(* IEC 61131-3 sources: daoli-st-library/DL_MathData (part 32) *)

(* ---- FC_DL_RangeOverlapCheck.st ---- *)
(*==============================================================================
 * 组件名称 (Component)  : FC_DL_RangeOverlapCheck
 * 所属子库 (Sublibrary) : DL_MathData
 * 当前版本 (Version)    : 1.0.0
 * 分类     (Category)   : 区间关系判定函数（Function · Comparator / Pure function）
 * 兼容性   (Platform)   : CODESYS 3.5 / TwinCAT 3 / 汇川 InoProShop / Machine Expert
 *                         仅依赖 Standard.library（ABS / MIN / MAX），零厂商方言
 * 功能描述 (Function)   : 判定两个实数区间 A、B 的几何关系（相离 / 仅端点相接 /
 *                         部分重叠 / 一方包含另一方 / 完全相等），并输出重叠长度。
 *                         输入是 4 个端点而非 1 个测量值，返回值为关系枚举，全程
 *                         无内部状态，可任意频次调用。用于配方参数域校验、时间窗
 *                         互斥检查、公差带叠加分析、安全包络与工艺窗口对撞检查。
 *
 * 【引脚契约 / Pin contract】
 *   输入 fA1        : REAL — 区间 A 端点 1 [任意工程单位]，无序自动对调；
 *   输入 fA2        : REAL — 区间 A 端点 2，同上；
 *   输入 fB1        : REAL — 区间 B 端点 1，无序自动对调；
 *   输入 fB2        : REAL — 区间 B 端点 2，同上；
 *   输入 bIncA      : BOOL — A 是否闭区间（含端点），默认 TRUE；
 *   输入 bIncB      : BOOL — B 是否闭区间，默认 TRUE；
 *   输出 fOverlapSpan : REAL — 重叠长度 [与输入同单位]，无重叠 = 0.0，恒非负；
 *   输出 bTouching    : BOOL — 仅端点相接（重叠长度 0 但边界重合）；
 *   输出 bValid       : BOOL — 四个输入全部有限（非 NaN、非无穷）= TRUE；
 *   输出 uErrorId     : UDINT — 事件码，0 = 无。本件全部码为信息级。
 *   返回  值          : E_DL_RangeRelation — 区间关系枚举，见下方成员语义表。
 *
 * 【关系枚举语义 / Relation enum semantics（同文件发布）】
 *   eInvalid  = 0  — 输入含非有限值（NaN / 无穷），关系不可判，重叠长度 0.0；
 *   eDisjoint = 10 — 完全相离（两区间之间有正间隙）；
 *   eTouching = 20 — 仅端点相接，重叠长度 0.0，bTouching 置位；
 *   ePartial  = 30 — 部分重叠（互相不包含，重叠长度大于 0）；
 *   eContains = 40 — 一方包含另一方（含端点恰好重合的包含）；
 *   eEqual    = 50 — 两端点均在容差内相等，重叠长度 = 区间长度。
 *
 * 【判定次序 / Decision order（写死，避免多解）】
 *   ① 有限性闸门 → 全部有限才继续，否则返回 eInvalid 并置 0121；
 *   ② 端点归一 → 每个区间内部排序，保证「下限 <= 上限」；
 *   ③ 相等判定 → 两端点同时落在容差内即 eEqual（先判，避免被包含分支吞掉）；
 *   ④ 相离判定 → 任一侧上限严格小于对侧下限减去容差，即 eDisjoint；
 *   ⑤ 相接判定 → 任一侧上限与对侧下限重合（容差内），即 eTouching；
 *   ⑥ 包含判定 → 一侧下限不大于对侧下限且上限不小于对侧上限，即 eContains；
 *   ⑦ 其余 → ePartial（此时重叠长度必然大于 0，无需再判）。
 *   次序不可调换：相等必须先于包含，相离必须先于相接，相接必须先于部分重叠。
 *
 * 【开闭区间口径 / Open and closed intervals（防误解声明）】
 *   ① 几何关系与开闭无关：「相接」只描述两组端点几何重合，开区间同样判相接；
 *   ② 开闭只影响「相接处那一个点是否属于公共交集」，其判据为
 *      bTouching AND bIncA AND bIncB —— 调用方按此合成，本件不额外输出第三态；
 *   ③ 部分重叠与包含的重叠长度按端点差值计算，不做「开区间减去两个端点」的
 *      离散化折算：连续量工程口径下端点测度为零，减去端点会引入 1 个单位误差；
 *   ④ 相等判定用容差而非判等（浮点判等红线）：两端点差值绝对值均小于容差即认为
 *      相等，容差取 1.0E-6，对应工程上「不可分辨」的量级。
 *
 * 【数值安全 / Numeric safety】
 *   N1 非有限值用「区间比较取反」识别：NaN 参与任何有序比较均为假，
 *      故 NOT(下限比较 AND 上限比较) 同时覆盖 NaN 与正负无穷，无需判等；
 *   N2 重叠长度在返回前置零下限保护：极少数退化输入可能算出负零附近的微小负值，
 *      一律钳到 0.0，保证输出恒非负（下游可直接做累加不打补丁）；
 *   N3 全件无除法、无开方、无累加迭代，不存在除零与溢出风险；
 *   N4 全件无循环、无数组访问，不存在越界风险。
 *
 * 【边界防错清单 / Boundary guard list】
 *   B1 输入非有限 → bValid FALSE、返回 eInvalid、重叠长度 0.0、置 0121（信息级）；
 *   B2 端点无序（如 A = [10, 0]）→ 自动对调后按归一区间判定，不置任何码；
 *   B3 零长度区间（两端点相等）→ 合法输入，参与全部关系判定，不特殊对待；
 *   B4 相接与部分重叠的边界由容差分割：端点差值绝对值小于容差判相接，
 *      否则按下限比较判重叠，容差量级远小于工程分辨率，不会误判真实重叠；
 *   B5 包含判定允许端点恰好重合（A 包含 B 且共端点），此时关系为 eContains
 *      而非 eEqual（eEqual 要求两端点都相等，先判，语义不重叠）。
 *
 * 【与既有件的职责边界 / Family separation（本族唯一二元件）】
 *   FC_DL_LimitClassify    = 判单个测量值落在哪一档（单点 → 档位）；
 *   FC_DL_Hysteresis       = 判单个测量值的迟滞切换（单点 + 历史 → 开关）；
 *   FB_DL_ToleranceWindow  = 判单个测量值是否落在公差带（单点 → 布尔）；
 *   本件                   = 判两个区间之间的关系（四点 → 关系枚举），
 *   输入元数不同、返回类型不同，四者不可互相替代。
 *
 * 【调用示例 / Call example（仅行注释，不嵌套块注释）】
 *   // 配方切换前校验：新工艺窗口与安全包络是否相撞
 *   // eRel := FC_DL_RangeOverlapCheck(fA1 := fSafeLo, fA2 := fSafeHi,
 *   //        fB1 := fNewLo, fB2 := fNewHi, bIncA := TRUE, bIncB := TRUE,
 *   //        fOverlapSpan => fOverlap, bTouching => bTouch,
 *   //        bValid => bCfgValid, uErrorId => uRelErr);
 *   // IF eRel = E_DL_RangeRelation.ePartial OR eRel = E_DL_RangeRelation.eContains THEN
 *   //     bRejectRecipe := TRUE;
 *   // END_IF
 *
 * 【平台移植注意 / Porting notes】
 *   仅用 ABS / MIN / MAX 三个标准函数与有序比较，无舍入模式依赖；
 *   容差与有限性阈值全部来自 VAR CONSTANT，换平台无需改逻辑；
 *   返回枚举类型随本文件发布，导入顺序上本文件不依赖任何其他 DL_ 组件。
 *
 * 【工程背景与应用场景 / Background and use cases】
 *   ① 配方参数域校验：新配方允许的温度带与设备安全包络相撞时拒绝下发；
 *   ② 时间窗互斥检查：两班次的作业窗若部分重叠，提示排程冲突；
 *   ③ 公差带叠加：来料公差带与装配公差带仅端点相接时，判定为「临界合格」；
 *   ④ 安全包络对撞：机器人可达包络与围栏安全距离带的重叠长度用于风险评估。
 *
 * 【验收向量 / Acceptance vectors】
 *   V1 部分重叠：A = [0, 10]、B = [5, 15] → ePartial、重叠长度 5.0；
 *   V2 端点相接：A = [0, 10]、B = [10, 20] → eTouching、重叠长度 0.0、bTouching；
 *   V3 包含：A = [0, 10]、B = [2, 8] → eContains、重叠长度 6.0；
 *   V4 相离：A = [0, 10]、B = [20, 30] → eDisjoint、重叠长度 0.0；
 *   V5 相等：A = [0, 10]、B = [0, 10] → eEqual、重叠长度 10.0；
 *   V6 无序端点：A = [10, 0]、B = [5, 15] → 归一后同 V1，ePartial、5.0；
 *   V7 非有限：fA1 为 NaN → eInvalid、bValid FALSE、uErrorId 0121。
 *
 * 【事件码表 / Event code table（全部信息级，不置报警位）】
 *   16#0001_0121  输入含非有限值，关系不可判，返回 eInvalid 与重叠长度 0.0。
 *
 * 修订历史 (Revision)   :
 *   2026-11-15  v1.0.0  首版落盘（Round 11 · 泳道 A · LGF Comparator 组）
 *
 * 同文件发布类型 (Co-published type) : E_DL_RangeRelation（本函数返回枚举，
 *   按库内惯例随宿主 POU 同文件发布，禁止在其他文件重复声明同名枚举）。
 *============================================================================*)
TYPE E_DL_RangeRelation :
(
    eInvalid  := 0,    // 输入非有限值，关系不可判 / Inputs not finite, relation undecidable
    eDisjoint := 10,   // 完全相离，存在正间隙 / Fully disjoint with a positive gap
    eTouching := 20,   // 仅端点相接，重叠长度为零 / Endpoint touch only, zero overlap
    ePartial  := 30,   // 部分重叠，互不包含 / Partial overlap, neither contains the other
    eContains := 40,   // 一方包含另一方 / One range contains the other
    eEqual    := 50    // 两端点均在容差内相等 / Both endpoints equal within tolerance
);
END_TYPE

FUNCTION FC_DL_RangeOverlapCheck : E_DL_RangeRelation
VAR_INPUT
    fA1     : REAL;                        // 区间 A 端点 1 [工程单位]，无序自动对调 / Range A endpoint 1 [EU], auto-swapped
    fA2     : REAL;                        // 区间 A 端点 2 [工程单位] / Range A endpoint 2 [EU]
    fB1     : REAL;                        // 区间 B 端点 1 [工程单位]，无序自动对调 / Range B endpoint 1 [EU], auto-swapped
    fB2     : REAL;                        // 区间 B 端点 2 [工程单位] / Range B endpoint 2 [EU]
    bIncA   : BOOL := TRUE;                // A 是否闭区间，含端点 / A closed interval flag, endpoints included
    bIncB   : BOOL := TRUE;                // B 是否闭区间，含端点 / B closed interval flag, endpoints included
END_VAR
VAR_OUTPUT
    fOverlapSpan : REAL;                   // 重叠长度 [工程单位]，无重叠 0.0，恒非负 / Overlap length [EU], zero when none, never negative
    bTouching    : BOOL;                   // 仅端点相接（几何重合，与开闭无关）/ Endpoint touch only, independent of openness
    bValid       : BOOL;                   // 四个输入全为有限值 / All four inputs are finite
    uErrorId     : UDINT;                  // 事件码，0 = 无 / Event code, 0 = none
END_VAR
VAR
    _fLoA   : REAL;                        // 区间 A 归一下限 [工程单位] / Normalised lower bound of range A [EU]
    _fHiA   : REAL;                        // 区间 A 归一上限 [工程单位] / Normalised upper bound of range A [EU]
    _fLoB   : REAL;                        // 区间 B 归一下限 [工程单位] / Normalised lower bound of range B [EU]
    _fHiB   : REAL;                        // 区间 B 归一上限 [工程单位] / Normalised upper bound of range B [EU]
    _fTmp   : REAL;                        // 对调临时量 [工程单位] / Swap temporary [EU]
    _fLo    : REAL;                        // 重叠区间下限 = 两个下限的较大者 [工程单位] / Overlap lower bound, the larger of both [EU]
    _fHi    : REAL;                        // 重叠区间上限 = 两个上限的较小者 [工程单位] / Overlap upper bound, the smaller of both [EU]
    _bFinite : BOOL;                       // 有限性闸门标志 / Finiteness gate flag
END_VAR
VAR CONSTANT
    DL_FLOAT_EPS  : REAL  := 1.0E-6;       // 端点比较容差 [工程单位] / Endpoint comparison epsilon [EU]
    DL_INF_LIM    : REAL  := 1.0E37;       // 非有限值判据阈值，超此视为无穷 / Non-finite threshold, beyond is infinity
    DL_SPAN_ZERO  : REAL  := 0.0;          // 重叠长度下界，恒非负 / Overlap length lower bound, never negative
    DL_ERR_NONFIN : UDINT := 16#0001_0121; // 输入非有限值的信息级码 / Info code for non-finite inputs
END_VAR

(*------------------------------------------------------------------------------
 * 段 1｜返回值与输出预置（函数必须先给出安全返回值）
 *      Preset the return value and the outputs
 *   默认返回 eInvalid：任何早退路径都天然带着「不可判」语义，不会误报相离。
 *-----------------------------------------------------------------------------*)
FC_DL_RangeOverlapCheck := E_DL_RangeRelation.eInvalid;   // 返回值预置不可判（Return preset to undecidable）
fOverlapSpan := DL_SPAN_ZERO;              // 重叠长度预置 0（Overlap span preset to zero）
bTouching    := FALSE;                     // 相接标志预置（Touch flag preset）
bValid       := TRUE;                      // 有效性预置通过（Validity preset to pass）
uErrorId     := 16#0000_0000;              // 事件码预清零（Event code preset to zero）
_bFinite     := TRUE;                      // 有限性闸门预置通过（Finiteness gate preset to pass）

(*------------------------------------------------------------------------------
 * 段 2｜有限性闸门（边界 B1 / 数值安全 N1）
 *      Finiteness gate
 *   NaN 与任何有序比较的结果均为假，故「比较区间取反」同时覆盖 NaN 与无穷，
 *   不必使用浮点判等，也不依赖任何厂商的非有限值判定函数。
 *-----------------------------------------------------------------------------*)
IF NOT ((fA1 <= DL_INF_LIM) AND (fA1 >= -DL_INF_LIM)) THEN   // 端点 A1 非有限（A1 not finite）
    _bFinite := FALSE;                     // 闸门关闭（Close the gate）
END_IF
IF NOT ((fA2 <= DL_INF_LIM) AND (fA2 >= -DL_INF_LIM)) THEN   // 端点 A2 非有限（A2 not finite）
    _bFinite := FALSE;                     // 闸门关闭（Close the gate）
END_IF
IF NOT ((fB1 <= DL_INF_LIM) AND (fB1 >= -DL_INF_LIM)) THEN   // 端点 B1 非有限（B1 not finite）
    _bFinite := FALSE;                     // 闸门关闭（Close the gate）
END_IF
IF NOT ((fB2 <= DL_INF_LIM) AND (fB2 >= -DL_INF_LIM)) THEN   // 端点 B2 非有限（B2 not finite）
    _bFinite := FALSE;                     // 闸门关闭（Close the gate）
END_IF

IF NOT _bFinite THEN                       // 任一输入不可判（Any input undecidable）
    bValid   := FALSE;                     // 有效性置假（Validity cleared）
    uErrorId := DL_ERR_NONFIN;             // 置非有限值信息码（Raise the non-finite info code）
    RETURN;                                // 早退，返回值保持 eInvalid（Early exit, return stays eInvalid）
END_IF

(*------------------------------------------------------------------------------
 * 段 3｜端点归一（边界 B2：无序端点自动对调）
 *      Endpoint normalisation, unordered endpoints are swapped
 *   归一后不可能出现「下限大于上限」，后续全部比较都是同向比较。
 *-----------------------------------------------------------------------------*)
_fLoA := fA1;                              // A 下限暂存端点 1（A lower bound takes endpoint 1）
_fHiA := fA2;                              // A 上限暂存端点 2（A upper bound takes endpoint 2）
IF _fLoA > _fHiA THEN                      // 端点逆序（Endpoints in reverse order）
    _fTmp := _fLoA;                        // 暂存下限（Save the lower bound）
    _fLoA := _fHiA;                        // 下限取原上限（Lower takes the former upper）
    _fHiA := _fTmp;                        // 上限取原下限（Upper takes the former lower）
END_IF

_fLoB := fB1;                              // B 下限暂存端点 1（B lower bound takes endpoint 1）
_fHiB := fB2;                              // B 上限暂存端点 2（B upper bound takes endpoint 2）
IF _fLoB > _fHiB THEN                      // 端点逆序（Endpoints in reverse order）
    _fTmp := _fLoB;                        // 暂存下限（Save the lower bound）
    _fLoB := _fHiB;                        // 下限取原上限（Lower takes the former upper）
    _fHiB := _fTmp;                        // 上限取原下限（Upper takes the former lower）
END_IF

_fLo := MAX(_fLoA, _fLoB);                 // 重叠下限 = 两个下限的较大者（Overlap lower bound）
_fHi := MIN(_fHiA, _fHiB);                 // 重叠上限 = 两个上限的较小者（Overlap upper bound）

(*------------------------------------------------------------------------------
 * 段 4｜关系判定（判定次序写死：相等 → 相离 → 相接 → 包含 → 部分）
 *      Relation decision in the frozen order
 *   次序不可调换，理由见头注释「判定次序」段；每支都显式给出重叠长度。
 *-----------------------------------------------------------------------------*)
IF (ABS(_fHiA - _fHiB) < DL_FLOAT_EPS) AND (ABS(_fLoA - _fLoB) < DL_FLOAT_EPS) THEN
    FC_DL_RangeOverlapCheck := E_DL_RangeRelation.eEqual;   // 相等：两端点均在容差内（Both endpoints equal within epsilon）
    fOverlapSpan := _fHiA - _fLoA;         // 重叠长度 = 区间长度（Overlap equals the range length）
ELSIF (_fHiA < _fLoB - DL_FLOAT_EPS) OR (_fHiB < _fLoA - DL_FLOAT_EPS) THEN
    FC_DL_RangeOverlapCheck := E_DL_RangeRelation.eDisjoint; // 相离：存在正间隙（A positive gap exists）
    fOverlapSpan := DL_SPAN_ZERO;          // 相离无重叠（No overlap when disjoint）
ELSIF (ABS(_fHiA - _fLoB) < DL_FLOAT_EPS) OR (ABS(_fHiB - _fLoA) < DL_FLOAT_EPS) THEN
    FC_DL_RangeOverlapCheck := E_DL_RangeRelation.eTouching; // 相接：端点几何重合（Endpoints coincide geometrically）
    fOverlapSpan := DL_SPAN_ZERO;          // 相接重叠长度为零（Zero overlap on a touch）
    bTouching    := TRUE;                  // 置相接标志（Raise the touch flag）
ELSIF ((_fLoA <= _fLoB + DL_FLOAT_EPS) AND (_fHiA >= _fHiB - DL_FLOAT_EPS)) OR
      ((_fLoB <= _fLoA + DL_FLOAT_EPS) AND (_fHiB >= _fHiA - DL_FLOAT_EPS)) THEN
    FC_DL_RangeOverlapCheck := E_DL_RangeRelation.eContains; // 包含：一方完全覆盖另一方（One range covers the other）
    fOverlapSpan := _fHi - _fLo;           // 重叠长度 = 被包含区间的长度（Overlap equals the inner range length）
ELSE
    FC_DL_RangeOverlapCheck := E_DL_RangeRelation.ePartial; // 部分重叠：互不包含（Partial overlap, neither contains）
    fOverlapSpan := _fHi - _fLo;           // 重叠长度 = 交集长度（Overlap equals the intersection length）
END_IF

(*------------------------------------------------------------------------------
 * 段 5｜重叠长度非负保护（数值安全 N2）
 *      Non-negative guard of the overlap span
 *   浮点舍入可能让理论为零的交集算出极小的负值，一律钳到 0，
 *   保证下游可直接累加与比较，不必各自打补丁。
 *-----------------------------------------------------------------------------*)
IF fOverlapSpan < DL_SPAN_ZERO THEN        // 重叠长度出现负值（A negative span appeared）
    fOverlapSpan := DL_SPAN_ZERO;          // 钳到 0，维持非负承诺（Clamp to zero, keep the promise）
END_IF
END_FUNCTION

(* ---- FC_DL_StringFixedField.st ---- *)
(*==============================================================================
 * 组件名称 (Component)  : FC_DL_StringFixedField
 * 所属子库 (Sublibrary) : DL_MathData
 * 归属目录 (Directory)  : C:\Library\DL_MathData
 * 当前版本 (Version)    : 1.0.0
 * 分类/来源标签         : 函数（FUNCTION）· 纯函数 · 定宽字段填充与对齐
 *                         lgf-datahandling / fixed-field / r37-reference
 * 兼容性   (Platform)   : CODESYS 3.5 / TwinCAT 3 / 汇川 InoProShop / 施耐德
 *                         Machine Expert；仅用 Standard.library 的 LEN / MID /
 *                         CONCAT / MIN，字符串声明一律显式带长度
 * 功能一句话 (Summary)  : 把任意文本装进定宽字段（左对齐或右对齐、指定填充字符），
 *                         并在发生裁剪时显式置截断标志与事件码。
 *
 * 本件存在的意义 (Why this unit exists)：
 *   本件存在的意义是把 R37 变成可复制的写法。全库所有「往定长缓冲写串」的地方，
 *   都可以照本件的四步顺序抄：先算一次源长度，再与目标宽度比较，比较成立就先置
 *   截断标志与码，最后才写缓冲。顺序一旦颠倒（先 CONCAT 再回夹、或回夹时不置标志），
 *   现场就会出现「字段看着对、内容被砍了一半、日志里一个字都没有」的事故。
 *   本件是全库唯一一处必须在写入前预判长度的地方，因此写成了可当范本读的样子。
 *
 * 功能描述 (Function)   : 先校验宽度契约，再解析填充字符，然后一次取源长度并与宽度
 *                         比较，按允许与否决定「截断写出」或「拒绝构造」，最后用
 *                         CONCAT 把核心段与填充段拼成恰好 nWidth 个字符的字段。
 *                         典型现场用途：定长报文拼装（固定列宽协议）、CSV 列对齐、
 *                         HMI 固定列显示、条形码定长补位、打印模板的等宽排版。
 * 与既有件边界 (Boundary): FC_DL_StringTrim 去首尾空白、FC_DL_StringSplit 拆分、
 *                         FC_DL_StringReplaceAll 替换。三者都改变内容而不改宽度；
 *                         本件只改宽度与对齐，内容字符顺序不动（除裁剪尾部）。
 *                         宽度是契约参数，本件不猜、不钳、不补零。
 * 设计要点 (Key notes)  : ① 源长度只取一次（R38），其后所有比较与循环上界都用该副本；
 *                         ② 裁剪判定先于任何写入（R37），标志置位先于结果构造；
 *                         ③ 拼装只用 CONCAT 与单字符填充，绝不用取子串的函数去「凑宽度」，
 *                           也不做「先拼后夹」的回夹写法；
 *                         ④ 出口长度天然等于宽度（核心段加填充段恰好补齐），总长不超过
 *                           声明上限，故不存在赋值时的静默截断；
 *                         ⑤ 每次进入先把结果清空，杜绝上一次调用的残留字符。
 *                         ⑥ 纯函数：无内部状态、无跨周期残留，同入参同结果。
 *
 * 【R37 四步顺序（本件样板，调用方照抄即可）】
 *   第 1 步  nSrcLen := LEN(sValue)                         只取一次，锁存
 *   第 2 步  IF nSrcLen > MIN(nWidth, DL_SFF_MAXLEN) THEN  与目标宽度比较（宽度与上限取小）
 *   第 3 步      bTruncated := TRUE                          先置标志，先于任何写入
 *   第 4 步      按 bAllowTrunc 决定截断写出还是拒绝构造     最后才写缓冲
 *
 * 【验收向量 / Acceptance vectors】
 *   V1  源「ABC」、宽度 6、左对齐 → 字段「ABC 加三个空格」、写出 6、不截断
 *   V2  源「ABC」、宽度 6、右对齐 → 字段「三个空格加 ABC」、写出 6
 *   V3  V-B 主向量（R37 核心）：源「ABCDEFGHIJ」、宽度 5、允许截断
 *       → 字段「ABCDE」、截断标志为真、码 0147；裁剪发生必须有人报警
 *   V4  V-B 拒绝路：同源同宽、不允许截断 → 返回假、字段空串、写出 0、码 0148、
 *       截断标志仍为真（事实发生了，只是没写出去）
 *   V5  V-A 域外：宽度 0 或宽度 300 → 返回假、码 0224；宽度不钳位，
 *       因为宽度是契约，猜不得
 *   V6  残留专测：连续两次调用，第二次源为空串 → 字段必须是纯填充，不残留上次内容
 *   V7  V-D 填充字符纠正：填充串为空 → 退回空格并置 0149，字段仍按宽度构造
 *
 * 开源溯源 (Origin)     : 来源标签 lgf-datahandling。LGF（Libre Graphical Framework）
 *                         为免费闭源发布的公开函数库手册，本件仅借鉴其数据处理组
 *                         「定长字段填充与对齐」这一功能分类的存在性，以及「源、宽度、
 *                         填充字符、对齐方式」四参数域的组织方式；许可证按其发布方
 *                         条款仅作分类参考，本件零代码行、零注释、零数据结构引用，
 *                         属 clean-room 独立实现，不构成衍生作品。
 * 码位说明 (Codes)      : 信息 16#0001_0147 已按允许截断 ｜ 16#0001_0148 已拒绝构造
 *                         16#0001_0149 填充串长度已纠正
 *                         故障 16#0001_0224 宽度域外。取号见本轮规格 §3.2。
 *                         码位优先级：0224 最高，其次 0148，再次 0147，最后 0149。
 * 依赖说明 (Depends)    : 无 DL_ 内部依赖；仅 Standard.library 的 LEN / MID / CONCAT / MIN。
 * 镜像量清单 (R38)      : nSrcLen 是本件唯一的锁存量，入口一次导出；唯一消费点集中在
 *                         段 4 的比较与段 5 的核心段构造两处，两处读的都是同一个副本，
 *                         全文不再对入参串取长度。
 * 偏离留档 (Deviation)  : 形参的字符串长度用字面量 255 声明，逻辑区用常量
 *                         DL_SFF_MAXLEN 表达同一上界。原因：IEC 的类型声明不接受
 *                         本 POU 内声明的常量，两者必须字面一致，此处已对齐并在
 *                         依赖说明中标注，不构成双源。
 * 红线自检 (Redline)    : 零全局变量表依赖 ｜ 零外部变量声明 ｜ 零物理地址直写
 *                         纯 IEC 61131-3 ｜ 无除法故无除零面 ｜ 循环上界由已钳位标量给定
 *                         全变量双语同行注释 ｜ 状态机 N/A（纯函数）｜ 无定时器实例
 * 修订历史 (Revision)   : 2026-11-15  v1.0.0  首版入库（Round 13 · 泳道 B 定长串族收口）
 *============================================================================*)

(*==============================================================================
 * 拼装示意 (Assembly geometry)，以源「ABC」、宽度 6 为例：
 *   核心段「ABC」长 3，填充段长 6 减 3 等于 3
 *   左对齐：核心段在前，结果为「ABC」加三个填充字符
 *   右对齐：填充段在前，结果为三个填充字符加「ABC」
 *   两者长度都恰好 6，不需要任何回夹，也就不存在「回夹了但没人知道」的面
 *   若源长 10、宽度 5：核心段按字符逐个取前 5 个，裁剪标志在此之前已置真
 *============================================================================*)

FUNCTION FC_DL_StringFixedField : BOOL
VAR_INPUT
    sValue      : STRING(255);      // 源文本 [ASCII]，定长 255 / Source text, fixed 255 characters
    nWidth      : INT;              // 目标字段宽度 [字符]，域 1 到 255，域外直接拒绝 / Target field width, 1 to 255, rejected outside
    sPad        : STRING(1) := ' '; // 填充字符，只取首字符 [字符] / Pad character, only the first character is used
    bAlignRight : BOOL := FALSE;    // 对齐方式，真为右对齐（左补），默认为左对齐 / TRUE right aligns, FALSE left aligns
    bAllowTrunc : BOOL := FALSE;    // 允许截断，真则裁剪写出，假则拒绝构造 / TRUE truncates and writes, FALSE refuses
END_VAR
VAR_OUTPUT
    sField      : STRING(255);      // 定宽字段结果 [ASCII]，成功时长度恰为宽度 / Fixed width field, exactly the width on success
    bTruncated  : BOOL;             // 是否发生裁剪，裁剪发生时必须为真 / Set true whenever truncation happened
    nWritten    : INT;              // 实际字段长度 [字符]，域 0 到 255 / Field length written, 0 to 255
    uErrorId    : UDINT;            // 事件码，0 表示无事件 / Event code, zero means none
END_VAR
VAR
    sPadChar  : STRING(1);   // 生效填充字符，单字符 [字符] / Effective pad character
    sCore     : STRING(255); // 核心段，裁剪后长度不超过宽度 [ASCII] / Core segment, never longer than the width
    sRun      : STRING(255); // 填充段，长度等于宽度减核心段长 [ASCII] / Pad run, width minus core length
    nSrcLen   : INT;         // 锁存的源文本长度 [字符]，全件唯一消费点 / Latched source length, the single source of truth
    nUse      : INT;         // 核心段实际取用长度 [字符] / Core segment length actually used
    nFill     : INT;         // 填充字符个数 [个] / Number of pad characters
    nPadLen   : INT;         // 填充串声明的实际长度 [字符] / Actual length of the pad string
    nI        : INT;         // 字符构造循环下标 [索引] / Character build loop index
    uCode     : UDINT;       // 码位暂存，出口单点写入 [码] / Code staging, written once at the exit
END_VAR
VAR CONSTANT
    DL_SFF_MAXLEN : INT := 255;   // 定长上限 [字符]，与形参声明一致 / Fixed length limit, matches the declarations
    DL_SFF_ONE    : INT := 1;     // 单字符长度参数 [字符] / Single character length argument
END_VAR

(*------------------------------------------------------------------------------
 * 段 1｜输出预置与残留清除（边界 B1）：结果先清空，杜绝上一次调用的残留字符
 *      Pre-set and clear: the field is emptied so nothing from the previous call survives
 *      这一步必须排在所有分支之前，否则「拒绝构造」路径会露出上一次的旧字段
 *      This must run before any branch, otherwise the refusal path leaks the old field
 *-----------------------------------------------------------------------------*)
FC_DL_StringFixedField := FALSE;
sField      := '';
sCore       := '';
sRun        := '';
sPadChar    := ' ';
bTruncated  := FALSE;
nWritten    := 0;
uErrorId    := 16#0000_0000;
uCode       := 16#0000_0000;
nSrcLen     := 0;
nUse        := 0;
nFill       := 0;
nPadLen     := 0;

(*------------------------------------------------------------------------------
 * 段 2｜宽度闸门（边界 B2）：宽度是契约参数，域外直接拒绝，绝不钳位
 *      Width gate: the width is a contract value, values outside the domain are refused
 *      钳位在这里是最坏的处理方式：调用方以为拿了 5 宽，实际拿到 255 宽，
 *      定长报文的列位会整体后移，且没有任何一条日志能对得上
 *      Clamping would shift every following column of a fixed layout report
 *-----------------------------------------------------------------------------*)
IF (nWidth < 1) OR (nWidth > DL_SFF_MAXLEN) THEN
    uErrorId := 16#0001_0224;   // 故障级：宽度域外，字段保持空串、写出 0
    RETURN;
END_IF

(*------------------------------------------------------------------------------
 * 段 3｜填充字符解析（边界 B3）：只取首字符，空串退回空格并报纠正码
 *      Pad resolution: take the first character only, an empty pad falls back to a space
 *-----------------------------------------------------------------------------*)
nPadLen := LEN(sPad);
IF nPadLen >= DL_SFF_ONE THEN
    sPadChar := MID(sPad, DL_SFF_ONE, DL_SFF_ONE);   // 位置 1 起取一个字符 / One character starting at position one
    IF nPadLen <> DL_SFF_ONE THEN
        uCode := 16#0001_0149;   // 信息级：填充串长度不是 1，已取首字符
    END_IF
ELSE
    sPadChar := ' ';             // 空填充串：退回空格，字符本身仍合法
    uCode    := 16#0001_0149;
END_IF

(*------------------------------------------------------------------------------
 * 段 4｜源长度一次锁存与裁剪预判（边界 B4，R37 主战场）：先判后写，标志先行
 *      Latch the source length and pre-judge truncation: judge first, flag first
 *      四步顺序不可颠倒：取长度、比较、置标志、再决定写出或拒绝
 *      The four steps are order critical, a reordered version loses the evidence
 *-----------------------------------------------------------------------------*)
nSrcLen := LEN(sValue);
IF nSrcLen < 0 THEN
    nSrcLen := 0;
END_IF

(* 裁剪门限双保险：字段宽度与声明上限同时参与，两者的较小者才是界
 * Double bounded: the smaller of the field width and the declared limit is the bound
 * 宽度已在段 2 限制在 1 到 255，故此处两界等价，写法上把「比长度」这件事显式化 *)
IF nSrcLen > MIN(nWidth, DL_SFF_MAXLEN) THEN

    bTruncated := TRUE;          // 第 3 步：事实先记录，早于任何写入

    IF NOT bAllowTrunc THEN
        (* 第 4 步之拒绝路：不构造字段，把决定权交回调用方 *)
        (* Refusal path: build nothing and leave the decision to the caller *)
        uErrorId := 16#0001_0148;
        RETURN;                  // 字段保持空串，写出保持 0
    END_IF

    uCode := 16#0001_0147;       // 第 4 步之裁剪路：允许截断，码位优先于填充纠正码
    nUse  := nWidth;

ELSE

    nUse := nSrcLen;             // 源不超宽，核心段全取 / The source fits, the whole text is the core

END_IF

(*------------------------------------------------------------------------------
 * 段 5｜核心段构造（边界 B5）：未裁剪直取，裁剪时逐字符取前 nUse 个
 *      Core segment build: assign directly when short enough, else copy character by character
 *      逐个字符取而不是对源取子串后回夹：路径唯一，长度由循环次数决定，
 *      既不依赖平台的子串边界行为，也不会出现「夹了但没报」的第二种写法
 *      Copying per character keeps the length structurally equal to the loop bound
 *-----------------------------------------------------------------------------*)
IF nUse >= nSrcLen THEN
    sCore := sValue;
ELSE
    FOR nI := 1 TO nUse DO
        sCore := CONCAT(sCore, MID(sValue, DL_SFF_ONE, nI));
    END_FOR;
END_IF

(*------------------------------------------------------------------------------
 * 段 6｜填充段构造（边界 B6）：个数由宽度减核心段长决定，恒非负
 *      Pad run build: the count is width minus core length, always non-negative
 *      nUse 最大等于 nWidth，故 nFill 最小为 0，循环上界天然合法
 *-----------------------------------------------------------------------------*)
nFill := nWidth - nUse;
IF nFill < 0 THEN
    nFill := 0;                  // 结构性保证已成立，仍显式兜底
END_IF

FOR nI := 1 TO nFill DO
    sRun := CONCAT(sRun, sPadChar);
END_FOR;

(*------------------------------------------------------------------------------
 * 段 7｜拼装与出口（边界 B7）：总长恰为宽度，赋值不存在静默截断
 *      Assembly and exit: the total length equals the width, no silent truncation
 *      核心段长加填充段长恒等于宽度，且宽度已限制在 255 以内
 *      Core plus pad always equals the width, which is already bounded by 255
 *-----------------------------------------------------------------------------*)
IF bAlignRight THEN
    sField := CONCAT(sRun, sCore);
ELSE
    sField := CONCAT(sCore, sRun);
END_IF

nWritten := MIN(nWidth, DL_SFF_MAXLEN);
uErrorId := uCode;               // 码位单点写入，全拍只写一次 / Single write point for the code
FC_DL_StringFixedField := TRUE;
END_FUNCTION

(* ---- FC_DL_StringToLReal.st ---- *)
(*==============================================================================
 * 组件名称 (Component)  : FC_DL_StringToLReal
 * 所属子库 (Sublibrary) : DL_MathData
 * 归属目录 (Directory)  : C:\Library\DL_MathData
 * 当前版本 (Version)    : 1.0.0
 * 分类/来源标签         : 函数（FUNCTION）· 纯函数 · 带校验的数值解析
 *                         lgf-datahandling / string-parse / validated-conversion
 * 兼容性   (Platform)   : CODESYS 3.5 / TwinCAT 3 / 汇川 InoProShop / 施耐德
 *                         Machine Expert；仅用 Standard.library 的 LEN / MID /
 *                         FIND / LIMIT / MIN / MAX，无厂商串转换函数依赖
 * 功能一句话 (Summary)  : 把定长 ASCII 文本严格解析成 LREAL，逐字符推进，拒绝一切
 *                         可疑输入，并报出首个非法字符的位置。
 * 功能描述 (Function)   : 语法为「可选符号、整数部、可选小数部、可选指数部」。解析
 *                         过程不调用平台的隐式串转数值功能，全部字符自行判定与推进，
 *                         因此三重收益：① 非法输入的行为在三家平台上完全一致；
 *                         ② 出错时能回答「错在第几个字符」，而不是只给一个零；
 *                         ③ 前缀合法、尾部夹脏字符时仍给出前缀值，方便现场判断是
 *                         报文截断还是字段串位。典型现场用途：条码与二维码文本入库、
 *                         CSV 报文列解析、HMI 手输设定值校验、第三方仪表 ASCII 应答
 *                         的数值字段提取。
 * 为什么自带解析 (Why)  : 三家平台对「字符串转实数」的非法输入行为不一致：有的返回
 *                         零、有的抛异常、有的静默截断，且都不告诉调用方错在第几位。
 *                         现场最贵的不是「转换失败」，而是「转换成功了但值不对」。
 * 与既有件边界 (Boundary): FC_DL_HexStringToBytes 处理十六进制到字节；本件处理十进制
 *                         文本到实数。二者共用「逐字符判定、失败保留前缀信息」的
 *                         口径，但字符集与输出类型完全不同，不重叠。
 * 设计要点 (Key notes)  : ① 长度一次锁存：入口取 LEN 存成局部量，其后所有循环上界、
 *                           下标判断、消费计数全部取自该副本，全文不再读入参长度；
 *                         ② 逐字符推进，不用任何回夹写法拼结果，也不靠平台转换函数；
 *                         ③ 先用状态推进做完语法判定，再统一做数值定稿，因此「语法
 *                           错误」与「数值越界」两类事件不会互相覆盖；
 *                         ④ 出口夹域：无论成功失败，fValue 一定落在调用方给定的
 *                           上下限之间，绝不输出无穷或非数；
 *                         ⑤ 纯函数：无内部状态、无跨周期残留，同入参同结果。
 *
 * 【解析状态映射表 / Parse phase map】
 *   起始态 0 期待符号、数字或小数点 ｜ 符号态 1 符号已取 ｜ 整数态 2 整数位推进
 *   小数态 3 小数位推进 ｜ 指数标记态 4 已见指数标记 ｜ 指数符号态 5 指数符号已取
 *   指数数字态 6 指数位推进。每个状态接受的输入集合在段 3 逐个分支写明，
 *   未列出的组合一律判非法字符，不存在「落到默认分支继续跑」的可能。
 *
 * 【验收向量 / Acceptance vectors】
 *   V1  文本「负号 1 2 点 5」→ 返回真、值 负 12.5、消费 5 字符、首错位 0
 *   V2  V-B 指数开关：文本「1 点 5 E 3」允许指数 → 1500.0；
 *       禁止指数 → 返回假、首错位 4、码 0144、值保留前缀 1.5
 *   V3  V-A 域外：文本「1 2 点 5 点 3」→ 返回假、码 0222、首错位 5、消费 4 字符
 *   V4  V-B 上限：文本「1 E 4 0」→ 返回假、码 0146、值夹到上限 1.0E30（不输出无穷）
 *   V5  V-C 锁存专测（R38）：调用方在本件返回后立即改写文本缓冲，本件内部所有边界
 *       都来自入口锁存的长度，结果不受影响；纯函数天然满足，此处作为纪律声明
 *   V6  V-D 出口夹域：文本「1 E 3 0」且上限 100 → 返回真、值 100.0、码 0145
 *   V7  全空白文本 → 返回假、码 0143、消费 0 字符、值 0.0
 *
 * 开源溯源 (Origin)     : 来源标签 lgf-datahandling。LGF（Libre Graphical Framework）
 *                         为免费闭源发布的公开函数库手册，本件仅借鉴其数据处理组
 *                         「字符串与数值互转按类型分函数、单一职责」的组织方式，以及
 *                         「带校验的转换器」这一功能分类的存在性；许可证按其发布方
 *                         条款仅作分类参考，本件零代码行、零注释、零数据结构引用，
 *                         属 clean-room 独立实现，不构成衍生作品。
 * 码位说明 (Codes)      : 信息 16#0001_0143 空或无有效数字 ｜ 16#0001_0144 尾随非法字符
 *                         16#0001_0145 结果已夹域 ｜ 16#0001_0146 指数超出保护域
 *                         故障 16#0001_0222 小数点重复 ｜ 16#0001_0223 结果非有限。
 *                         取号见本轮规格 §3.2，与 CRC8 子族 0141 到 0142 不重叠。
 * 依赖说明 (Depends)    : 无 DL_ 内部依赖；仅 Standard.library 的 LEN / MID / FIND /
 *                         LIMIT / MIN / MAX 与 INT_TO_LREAL 显式转换。
 * 镜像量清单 (R38)      : nLen 是本件唯一的锁存量，入口一次导出；唯一消费点集中在
 *                         段 2 的全空白预扫、段 3 的循环上界、段 5 的消费计数三处，
 *                         三处读的都是同一个局部副本，全文不再对入参串取长度。
 * 契约前置条件 (Contract): fMin 与 fMax 必须为有限值；两者倒置时按 MIN / MAX 自动
 *                         归正，不报错也不新增码位（上下限属组态参数，非运行数据）。
 * 偏离留档 (Deviation)  : 形参的字符串长度用字面量 40 声明，逻辑区用常量 DL_S2N_MAXLEN
 *                         表达同一上界。原因：IEC 的类型声明不接受本 POU 内声明的常量，
 *                         两者必须字面一致，此处已对齐，不构成双源。
 * 红线自检 (Redline)    : 零全局变量表依赖 ｜ 零外部变量声明 ｜ 零物理地址直写
 *                         纯 IEC 61131-3 ｜ 每处除法前判除数下限 ｜ 循环上界全常量化
 *                         全变量双语同行注释 ｜ 状态机 N/A（纯函数）｜ 无定时器实例
 * 修订历史 (Revision)   : 2026-11-15  v1.0.0  首版入库（Round 13 · 泳道 B 定长串族收口）
 *============================================================================*)

(*==============================================================================
 * 逐字符推演 (Character walk-through)，以「1 2 点 5 点 3」为例：
 *   第 1 字符 数字 1，由起始态进入整数态，尾数 1，有效位计数 1
 *   第 2 字符 数字 2，整数态继续，尾数 12，有效位计数 2
 *   第 3 字符 小数点，由整数态进入小数态，小数点计数 1
 *   第 4 字符 数字 5，小数态累加，尾数 125，小数位计数 1
 *   第 5 字符 小数点，当前已在小数态，小数点计数变 2，判定重复，停在第 5 位
 *   消费字符数为 4，首错位为 5，值按尾数 125 除以 10 得 12.5 保留
 *   若调用方只看返回值会以为「全错」，看值与位置才知道是小数点写了两遍
 *============================================================================*)

FUNCTION FC_DL_StringToLReal : BOOL
VAR_INPUT
    sText     : STRING(40);         // 待解析文本 [ASCII]，定长 40，冗余位填空格或空 / Text to parse, fixed length 40
    bAllowExp : BOOL := TRUE;       // 允许指数部，真则接受大写或小写 E / Allow the exponent part, both cases accepted
    fMin      : LREAL := -1.0E30;   // 输出下限 [工程单位]，越限钳位 / Lower clamp in engineering units
    fMax      : LREAL := 1.0E30;    // 输出上限 [工程单位]，越限钳位 / Upper clamp in engineering units
END_VAR
VAR_OUTPUT
    fValue    : LREAL;              // 解析结果 [工程单位]，失败时保留已解析前缀值 / Parsed value, keeps the parsed prefix on failure
    nCharUsed : INT;                // 已消费字符数 [个]，域 0 到 40 / Characters consumed, 0 to 40
    nBadPos   : INT;                // 首个非法字符位置 [位]，1 起，0 表示全部合法 / First invalid position, one based, zero when clean
    uErrorId  : UDINT;              // 事件码，0 表示无事件 / Event code, zero means none
END_VAR
VAR
    nLen        : INT;              // 锁存的文本有效长度 [字符]，全件唯一消费点 / Latched text length, the single source of truth
    nPos        : INT;              // 字符扫描下标 [位]，1 起 / Character scan index, one based
    nI          : INT;              // 通用循环下标，用于预扫与幂次循环 [索引] / Generic loop index for the pre-scan and power loop
    nState      : INT;              // 解析阶段号 [态]，取值含义见头注释映射表 / Parse phase number, see the map in the header
    sChar       : STRING(1);        // 当前字符，由标准 MID 取出 [字符] / Current character read with the standard MID
    nDigit      : INT;              // 当前字符的数字值 [数]，非数字为负 1 / Digit value of the current character, minus one when not a digit
    fMant       : LREAL;            // 尾数累加值，按十进制逐位左移再加 [无量纲] / Mantissa accumulator
    nSig        : INT;              // 已累加的有效数字位数 [个]，有上限保护 / Accumulated significant digits, capped
    nFrac       : INT;              // 已累加的小数位数 [个]，决定尺度分母 / Accumulated fractional digits, drives the scale divisor
    nExp        : INT;              // 指数绝对值累加 [无量纲]，最多取三位 / Exponent magnitude, at most three digits
    nExpDig     : INT;              // 已累加的指数位数 [个] / Accumulated exponent digit count
    nDotCnt     : INT;              // 小数点出现次数 [次]，用于重复判定 / Decimal point occurrences
    bSign       : BOOL;             // 尾数符号，真为负 / Mantissa sign, true means negative
    bExpSign    : BOOL;             // 指数符号，真为负 / Exponent sign, true means negative
    bOk         : BOOL;             // 语法与数值均通过标记 / Syntax and numeric checks passed
    bStop       : BOOL;             // 扫描停止标记，遇首个错误后置真 / Scan stop flag, set at the first error
    bAnyVisible : BOOL;             // 文本含至少一个非空白字符标记 / At least one non blank character present
    fDiv        : LREAL;            // 小数尺度分母 [无量纲] / Fractional scale divisor
    fPow        : LREAL;            // 指数幂次中间量 [无量纲] / Exponent power accumulator
    nAbsExp     : INT;              // 指数绝对值 [无量纲]，用于幂次循环次数 / Absolute exponent, drives the power loop
    fLo         : LREAL;            // 归一后的出口下限 [工程单位] / Normalised lower bound
    fHi         : LREAL;            // 归一后的出口上限 [工程单位] / Normalised upper bound
    uCode       : UDINT;            // 码位暂存，出口单点写入 [码] / Code staging, written once at the exit
END_VAR
VAR CONSTANT
    DL_S2N_MAXLEN  : INT := 40;                     // 文本长度上限 [字符]，与形参声明一致 / Text length limit, matches the declaration
    DL_S2N_SIGMAX  : INT := 18;                     // 有效数字累加上限 [位]，覆盖双精度可表示精度 / Significant digit cap
    DL_S2N_EXPMAX  : INT := 38;                     // 指数绝对值上限 [无量纲]，超出转保护域 / Exponent magnitude limit
    DL_S2N_TEN     : LREAL := 10.0;                 // 十进制基数 [无量纲] / Decimal radix
    DL_S2N_FINITE  : LREAL := 1.0E308;              // 有限性上界 [无量纲]，用于拦无穷与非数 / Finiteness bound
    DL_S2N_DIGITS  : STRING := '0123456789';        // 数字字符表，用 FIND 定位取数值 / Digit table queried with FIND
    DL_S2N_ST_START : INT := 0;                     // 起始态，期待符号、数字或小数点 / Start phase
    DL_S2N_ST_SIGN  : INT := 1;                     // 符号态，尾数符号已取 / Mantissa sign phase
    DL_S2N_ST_INT   : INT := 2;                     // 整数态，整数位推进 / Integer phase
    DL_S2N_ST_FRAC  : INT := 3;                     // 小数态，小数位推进 / Fraction phase
    DL_S2N_ST_E     : INT := 4;                     // 指数标记态，已见指数标记 / Exponent marker phase
    DL_S2N_ST_ESIGN : INT := 5;                     // 指数符号态，指数符号已取 / Exponent sign phase
    DL_S2N_ST_EDIG  : INT := 6;                     // 指数数字态，指数位推进 / Exponent digit phase
END_VAR

(*------------------------------------------------------------------------------
 * 段 1｜输出预置：值、消费数、首错位、码位全部先落确定值
 *      Pre-set the outputs so every exit path publishes a deterministic result
 *-----------------------------------------------------------------------------*)
FC_DL_StringToLReal := FALSE;
fValue      := 0.0;
nCharUsed   := 0;
nBadPos     := 0;
uErrorId    := 16#0000_0000;
uCode       := 16#0000_0000;
nState      := DL_S2N_ST_START;
sChar       := '';
nDigit      := -1;
fMant       := 0.0;
nSig        := 0;
nFrac       := 0;
nExp        := 0;
nExpDig     := 0;
nDotCnt     := 0;
bSign       := FALSE;
bExpSign    := FALSE;
bOk         := FALSE;
bStop       := FALSE;
bAnyVisible := FALSE;
fDiv        := 1.0;
fPow        := 1.0;
nLen        := 0;

(*------------------------------------------------------------------------------
 * 段 2｜长度一次锁存与空文本判定（边界 B1）
 *      Latch the length once and reject empty or blank-only text
 *      锁存后所有边界判断只用 nLen，不再读入参串，这是纪律不是偏好：
 *      分拍处理时入参可能被别的任务改写，混用两种来源会切出「有效但为空」的假段
 *      Every later boundary uses the latched copy only, never the live parameter
 *-----------------------------------------------------------------------------*)
nLen := LEN(sText);
IF nLen < 0 THEN
    nLen := 0;
ELSIF nLen > DL_S2N_MAXLEN THEN
    nLen := DL_S2N_MAXLEN;
END_IF

IF nLen = 0 THEN
    uErrorId := 16#0001_0143;   // 信息级：空文本，无有效数字
    RETURN;
END_IF

FOR nI := 1 TO nLen DO
    sChar := MID(sText, 1, nI);
    IF (sChar <> ' ') AND (sChar <> '$09') AND (sChar <> '$0D') AND (sChar <> '$0A') THEN
        bAnyVisible := TRUE;    // 见到任意非空白字符即可停止判定目的 / Any visible character clears the all blank case
    END_IF
END_FOR;

IF NOT bAnyVisible THEN
    uErrorId := 16#0001_0143;   // 信息级：全空白文本，与空文本同码
    RETURN;
END_IF

bOk := TRUE;   // 语法判定从真开始，逐字符推进，遇错置假 / Starts true, each character may clear it

(*------------------------------------------------------------------------------
 * 段 3｜逐字符推进（边界 B2/B3/B4）：字符分四类处理，非数字非符号非点全判非法
 *      Character walk: four classes handled, anything else is illegal
 *      顺序硬约束：先判小数点（它改变状态），再判数字（它可能刚进入状态），
 *      再判符号（只在起始或指数标记之后合法），最后兜底一切其它字符
 *      Order matters: point first, then digit, then sign, then the catch-all
 *-----------------------------------------------------------------------------*)
FOR nPos := 1 TO nLen DO

    IF NOT bStop THEN

        sChar  := MID(sText, 1, nPos);
        nDigit := FIND(DL_S2N_DIGITS, sChar) - 1;   // 命中为 0 到 9，未命中为负 1

        IF sChar = '.' THEN
            (* 小数点只允许出现在起始、符号后、整数部之后；在小数态再次出现即重复 *)
            (* A decimal point is legal at the start, after a sign, or once after the integer part *)
            IF (nState = DL_S2N_ST_START) OR (nState = DL_S2N_ST_SIGN) OR (nState = DL_S2N_ST_INT) THEN
                nState  := DL_S2N_ST_FRAC;
                nDotCnt := nDotCnt + 1;
            ELSIF nState = DL_S2N_ST_FRAC THEN
                nDotCnt  := nDotCnt + 1;
                bOk      := FALSE;
                bStop    := TRUE;
                nBadPos  := nPos;
                nCharUsed := nPos - 1;
                uCode    := 16#0001_0222;   // 故障级：小数点重复
            ELSE
                bOk      := FALSE;
                bStop    := TRUE;
                nBadPos  := nPos;
                nCharUsed := nPos - 1;
                uCode    := 16#0001_0144;   // 信息级：小数点出现在指数部
            END_IF

        ELSIF nDigit >= 0 THEN
            (* 数字在起始态或符号态出现，即进入整数部；在指数标记或指数符号后出现，进入指数数字态 *)
            (* A digit after the start or the sign opens the integer part, after a marker it opens the exponent *)
            IF (nState = DL_S2N_ST_START) OR (nState = DL_S2N_ST_SIGN) THEN
                nState := DL_S2N_ST_INT;
            ELSIF (nState = DL_S2N_ST_E) OR (nState = DL_S2N_ST_ESIGN) THEN
                nState := DL_S2N_ST_EDIG;
            END_IF

            IF nState = DL_S2N_ST_EDIG THEN
                IF nExpDig < 3 THEN
                    nExp    := nExp * 10 + nDigit;
                    nExpDig := nExpDig + 1;
                END_IF
            ELSE
                IF nSig < DL_S2N_SIGMAX THEN
                    fMant := fMant * DL_S2N_TEN + INT_TO_LREAL(nDigit);
                    nSig  := nSig + 1;
                    IF nState = DL_S2N_ST_FRAC THEN
                        nFrac := nFrac + 1;
                    END_IF
                END_IF
            END_IF

        ELSIF (sChar = '+') OR (sChar = '-') THEN
            (* 符号只在起始位置（尾数符号）或指数标记之后（指数符号）合法 *)
            (* A sign is legal only at the start or right after the exponent marker *)
            IF nState = DL_S2N_ST_START THEN
                bSign  := (sChar = '-');
                nState := DL_S2N_ST_SIGN;
            ELSIF nState = DL_S2N_ST_E THEN
                bExpSign := (sChar = '-');
                nState   := DL_S2N_ST_ESIGN;
            ELSE
                bOk      := FALSE;
                bStop    := TRUE;
                nBadPos  := nPos;
                nCharUsed := nPos - 1;
                uCode    := 16#0001_0144;   // 信息级：符号位置非法
            END_IF

        ELSIF (sChar = 'E') OR (sChar = 'e') THEN
            (* 指数标记只允许紧跟尾数，且必须由开关放行；未放行时按尾随非法字符处理 *)
            (* The marker must follow the mantissa and must be enabled, otherwise it counts as trailing garbage *)
            IF ((nState = DL_S2N_ST_INT) OR (nState = DL_S2N_ST_FRAC)) AND bAllowExp THEN
                nState := DL_S2N_ST_E;
            ELSE
                bOk      := FALSE;
                bStop    := TRUE;
                nBadPos  := nPos;
                nCharUsed := nPos - 1;
                uCode    := 16#0001_0144;
            END_IF

        ELSE
            (* 兜底：空格、制表、回车、换行、货币符号、千分位逗号等一律判非法 *)
            (* Catch-all: blanks, tabs, carriage returns, currency signs and thousands separators are illegal *)
            bOk      := FALSE;
            bStop    := TRUE;
            nBadPos  := nPos;
            nCharUsed := nPos - 1;
            uCode    := 16#0001_0144;
        END_IF

    END_IF

END_FOR;

(*------------------------------------------------------------------------------
 * 段 4｜终态校验（边界 B5）：必须收在整数态、小数态或指数数字态，且至少一位数字
 *      Final phase check: must end inside a digit bearing phase with at least one digit
 *      只有符号、只有小数点、只有指数标记这三种「半截输入」在此统一拦下
 *      Half finished inputs such as a lone sign or a lone point are stopped here
 *-----------------------------------------------------------------------------*)
IF bOk THEN
    (* 正向条件写成「非合法终态」，避免在合法分支里做无意义的自我赋值 *)
    (* Written as a negative test so the legal branch needs no self assignment *)
    IF NOT ((((nState = DL_S2N_ST_INT) OR (nState = DL_S2N_ST_FRAC)) AND (nSig > 0))
        OR ((nState = DL_S2N_ST_EDIG) AND (nExpDig > 0))) THEN
        bOk       := FALSE;
        nBadPos   := 0;
        nCharUsed := 0;
        uCode     := 16#0001_0143;   // 信息级：无完整数字
    ELSE
        nCharUsed := nLen;           // 全部字符合法消费 / Every character was legally consumed
    END_IF
END_IF

(*------------------------------------------------------------------------------
 * 段 5｜数值定稿（边界 B6/B7）：尺度、指数、符号三步依次作用，前缀值同样成立
 *      Numeric finalisation: scale, exponent and sign applied in that order
 *      语法失败时本段照跑：前缀值可能就是现场要的东西，丢掉它等于丢掉证据
 *      This stage runs even after a syntax error, the prefix value is evidence
 *-----------------------------------------------------------------------------*)
fValue := fMant;

fDiv := 1.0;
FOR nI := 1 TO nFrac DO
    fDiv := fDiv * DL_S2N_TEN;       // 分母最大 1.0E18，必然有限 / The divisor stays finite
END_FOR;
IF fDiv > 0.0 THEN
    fValue := fValue / fDiv;         // 判零后再除，除数恒不小于 1.0 / Guarded division, the divisor is at least one
END_IF

nAbsExp := nExp;   // 指数幅度：nExp 累加时只进正值，正负由 bExpSign 单独承担 / Magnitude only, the sign lives in bExpSign

IF nAbsExp > DL_S2N_EXPMAX THEN
    (* 指数超保护域：正向溢出落到有限极值，负向下溢落到零，两者都不输出无穷或非数 *)
    (* Exponent beyond the guard band: overflow lands on the finite bound, underflow on zero *)
    IF bExpSign THEN
        fValue := 0.0;               // 下溢：数值已小于可表示下限 / Underflow, the value collapsed
    ELSE
        fValue := DL_S2N_FINITE;     // 上溢：先落到有限上界 / Overflow, land on the finite bound
    END_IF
    IF uCode = 16#0000_0000 THEN
        uCode := 16#0001_0146;
    END_IF
    bOk := FALSE;
ELSIF nAbsExp > 0 THEN
    (* 指数在保护域内：正向做乘法，负向做判零后的除法，幂次循环上界不超过上限常量 *)
    (* Inside the guard band: multiply for a positive exponent, guarded divide for a negative one *)
    fPow := 1.0;
    FOR nI := 1 TO nAbsExp DO
        fPow := fPow * DL_S2N_TEN;
    END_FOR;
    IF bExpSign THEN
        IF fPow > 0.0 THEN
            fValue := fValue / fPow; // 判零后再除，除数恒不小于 10.0 / Guarded division, the divisor is at least ten
        END_IF
    ELSE
        fValue := fValue * fPow;
    END_IF
END_IF

IF bSign THEN
    fValue := -fValue;               // 符号最后作用，指数与尺度都不带符号 / The sign is applied last
END_IF

(* 有限性检查：两个比较同时成立才算有限，非数会让两个比较都为假，故此式一并拦截
 * Finiteness check: both comparisons must hold, a not-a-number fails both, so it is caught too *)
IF NOT ((fValue <= DL_S2N_FINITE) AND (fValue >= -DL_S2N_FINITE)) THEN
    bOk := FALSE;
    IF uCode = 16#0000_0000 THEN
        uCode := 16#0001_0223;       // 故障级：结果非有限
    END_IF
    fValue := 0.0;
END_IF

(*------------------------------------------------------------------------------
 * 段 6｜出口夹域（边界 B8，R43 精神）：值必须落在调用方给定区间内
 *      Exit clamp: the value always lands inside the caller supplied range
 *      上下限倒置时按 MIN / MAX 归正，组态笔误不应让输出跑到域外
 *      Inverted bounds are normalised with MIN and MAX, the output never leaves the domain
 *-----------------------------------------------------------------------------*)
fLo := MIN(fMin, fMax);
fHi := MAX(fMin, fMax);

IF fValue < fLo THEN
    fValue := fLo;
    IF uCode = 16#0000_0000 THEN
        uCode := 16#0001_0145;
    END_IF
ELSIF fValue > fHi THEN
    fValue := fHi;
    IF uCode = 16#0000_0000 THEN
        uCode := 16#0001_0145;
    END_IF
END_IF

(*------------------------------------------------------------------------------
 * 段 7｜码位单点写入与返回判定
 *      Single write point for the code and the return decision
 *      返回真仅限「语法通过且无码或仅夹域」；夹域后值仍可直接使用，故不判失败
 *      True only when the syntax passed and either no code or a clamp-only code
 *-----------------------------------------------------------------------------*)
uErrorId := uCode;
FC_DL_StringToLReal := bOk AND ((uCode = 16#0000_0000) OR (uCode = 16#0001_0145));
END_FUNCTION

(* ---- FC_DL_TempUnitConvert.st ---- *)
(*==============================================================================
 * 组件名称 (Component)  : FC_DL_TempUnitConvert
 * 所属子库 (Sublibrary) : DL_MathData
 * 当前版本 (Version)    : 1.0.1
 * 分类/来源标签         : lgf-converter（T2-1 LGF Converter 组回补）
 * 作者/日期             : Daoli Library / 2026-11-15
 * 兼容性   (Platform)   : CODESYS 3.5 / TwinCAT 3 / 汇川 InoProShop / Machine Expert
 *                         仅依赖 Standard.library（ABS），纯函数无状态
 * 功能简介 (Function)   : 摄氏 / 华氏 / 开尔文三温标两两互转。源 / 目标由枚举
 *                         单向选择（非 MODE 巨无霸：仅 3×3 查表映射，公式域固定）。
 *                         物理无效（低于绝对零度）置信息级诊断不阻断返回。
 *                         典型现场用途：热电阻 / 热电偶 HMI 显示单位切换、
 *                         进口设备华氏组态与国产摄氏台账的台账口径统一、
 *                         能耗报表开尔文热力学量换算。
 * 开源溯源 (Origin)     : 原创实现（参考 LGF 公开手册 Converter 分类中
 *                         温标换算族的功能分类与参数域），换算公式取自公开
 *                         温标定义，只借分类/参数域/命名，clean-room 实现，
 *                         未复制任何源码。来源标签：lgf-converter。
 * 依赖     (Depends)    : 无 DL_ 内部依赖；Standard.library: ABS
 *
 * 【接口契约 / Interface contract】
 *   返回值：换算结果 [目标温标单位]；枚举非法时恒为 0.0。
 *   输入  ：fVal 输入温度；eSrc 源温标；eDst 目标温标。
 *   输出  ：uErrorId 故障码（绝对零度信息级 / 枚举非法故障级）。
 *   纪律  ：纯函数同输入同输出；无内部状态；可安全放进 IF 表达式与
 *           多任务环境（无共享可变状态）。
 *
 * 【使用示例 / Usage example】
 *   VAR
 *       fShow : LREAL;      // HMI 显示值
 *       nErr  : UDINT;      // 诊断码
 *   END_VAR
 *   // 台账存摄氏，HMI 依用户语言显示华氏：
 *   fShow := FC_DL_TempUnitConvert(fVal := fLedger, eSrc := E_DL_TempUnit.eCelsius,
 *                                  eDst := E_DL_TempUnit.eFahrenheit,
 *                                  uErrorId => nErr);
 *   IF nErr = 16#0001_0110 THEN
 *       // 信息级：源值低于绝对零度，坏值溯源（如热电偶断线负满量程）
 *   END_IF
 *
 * 【设计决策：枚举对而非模式码 / Enum pair instead of a mode code】
 *   3×3 组合用"源枚举 + 目标枚举"两个引脚表达，取代单引脚 MODE 巨无霸
 *   （单模式码要为 9 条路径编 9 个号，组态可读性差且易填错号）。
 *   枚举对 + 单向基准链（先归一到摄氏）使公式域固定为 4 条，
 *   新增温标只需扩归一段与展开段各一个 CASE 分支。
 *
 * 【换算公式域 / Formula domain（公开温标定义）】
 *   K → C : C = K - 273.15        ｜ C → K : K = C + 273.15
 *   F → C : C = (F - 32) × 5 / 9  ｜ C → F : F = C × 9 / 5 + 32
 *   全部 9 条路径（含同标直通）都由这 4 条公式 + 直通覆盖，无组合爆炸。
 *
 * 【诊断链设计 / Diagnostic chain design】
 *   绝对零度诊断置信息级不阻断：断线 / 短路的模拟量常表现为负满量程
 *   （约 -327 度摄氏口径），截断为绝对零度会抹掉故障证据；
 *   照算输出让上层诊断链能看到"多不可能"，溯源更直接。
 *
 * 验收向量 (Acceptance) :
 *   V1 fVal = 100.0, eCelsius → eKelvin     ：返回 373.15（沸点）
 *   V2 fVal = 100.0, eCelsius → eFahrenheit ：返回 212.0（沸点华氏）
 *   V3 fVal =  32.0, eFahrenheit → eCelsius ：返回 0.0（冰点）
 *   V4 fVal = 300.0, eKelvin → eCelsius     ：返回 26.85（常温）
 *   V5 fVal = -40.0, eCelsius → eFahrenheit ：返回 -40.0（双温标交点）
 *
 * 【同标直通与往返一致性推演 / Pass-through and round-trip checks】
 *   P1 eCelsius → eCelsius, fVal = 23.4 → 返回 23.4（同标直通零损耗）
 *   P2 eKelvin → eKelvin,    fVal = 0.0 → 返回 0.0 且不置绝对零度诊断
 *      （0 K 恰为绝对零度，容差含等号口径，合法物理下界）
 *   P3 V5 往返：-40 F → C 得 -40.0，再 C → F 仍得 -40.0（交点往返零漂移）
 *   P4 V1 往返：373.15 K → C 得 100.0，再 C → K 仍得 373.15
 *      （单向基准链 + 双精度浮点，往返误差在 1E-9 容差内）
 *
 * 【拒绝路径推演 / Rejection path walk-through】
 *   R1 eSrc = 200（非法枚举）→ uErrorId=0001_0207、返回 0.0（B2）
 *   R2 eDst = 99（非法枚举） → uErrorId=0001_0208、返回 0.0（B2）
 *   R3 fVal = -300（摄氏，低于绝对零度）→ uErrorId=0001_0110 信息级，
 *      返回值照算（华氏口径 -452.0）不截断（B3 诊断链留证）
 *
 * 【调用开销与部署建议 / Cost and deployment notes】
 *   每次调用固定成本：至多两次乘除、一次加减与一个 CASE 分支，
 *   无循环无状态，可放心放进 HMI 刷新链与报表计算链高频调用；
 *   台账口径建议全程统一摄氏存储、显示层换算，
 *   避免多级换算叠加放大舍入误差。
 * 故障码表 (Error codes):
 *   16#0001_0110  归一后温度低于绝对零度（信息级，不阻断，返回值照算输出，
 *                 便于诊断链追溯坏值来源）
 *   16#0001_0207  源温标枚举非法（故障级，返回 0.0）
 *   16#0001_0208  目标温标枚举非法（故障级，返回 0.0）
 *   【码位终审】原拟 0004_0101 / 0004_0201 / 0004_0202 经全库复核冲突：0004
 *   段属 DL_Motion（公约 0.7 段位表），且三码已分别被 FB_DL_SingleAxis
 *   （0004_0101 指令丢弃、0004_0201 非法态、0004_0202 软限位越界）、
 *   FB_DL_AxisRelativeMove / FB_DL_AxisVelocityMove（0004_0201）占用。
 *   本体属 DL_MathData，已顺延至 0001_0110 / 0001_0207 / 0001_0208（无冲突）。
 * 红线自检 (Redline)    : R1 ✓ 零全局存储 / 零外部变量引用 ｜ R2 ✓ 零物理地址直写
 *                         R3 ✓ 纯 IEC 61131-3 ｜ R4 ✓ 枚举越界拒绝 + 绝对零度诊断 + 除数常量判零守卫
 *                         R5 ✓ 全变量与枚举项中英双语同行注释 ｜ R6 ✓ 纯函数无状态（R6 状态机 N/A）
 *                         R7 ✓ 无定时器 / 边沿实例（R7 N/A）
 * 边界契约 (Boundaries):
 *   B1 换算基准链：一律先归一到摄氏（K → C 减绝对零度偏移；F → C 按公开
 *      温标定义式），再从摄氏到目标；同标转换直通。
 *      单向基准链保证 3×3 = 9 条路径只用 4 个公式，公式域固定无组合爆炸。
 *   B2 枚举越界值（非 0/1/2）→ 置故障级码并返回 0.0：静默返回错误温标数值
 *      比返回 0 更危险（0 摄氏度与 0 开尔文差 273.15，工艺员一眼可辨）。
 *   B3 归一后低于绝对零度 → 置信息级码，返回值照算输出不截断，
 *      供诊断链追溯（如热电偶断线负满量程）。
 *   B4 纯函数：同输入同输出，无内部状态、无副作用，可安全放进 IF 表达式。
 * 修订历史 (Revision)   :
 *   2026-11-15  v1.0.0  首版落盘（Round 09 · 泳道 A · Level 0 原子族回补）
 *   2026-11-15  v1.0.1  终审修复：故障码 0004_0101 / 0004_0201 / 0004_0202 属
 *                       DL_Motion 段位且与 SingleAxis / AxisRelativeMove /
 *                       AxisVelocityMove 冲突，改归 DL_MathData 段
 *                       0001_0110 / 0001_0207 / 0001_0208，换算与返回语义零改动
 *============================================================================*)
TYPE E_DL_TempUnit :
(
    eCelsius    := 0,  // 摄氏度 [deg C] / Celsius
    eFahrenheit := 1,  // 华氏度 [deg F] / Fahrenheit
    eKelvin     := 2   // 开尔文 [K] / Kelvin
);
END_TYPE

FUNCTION FC_DL_TempUnitConvert : LREAL    // 返回换算结果 [目标温标单位] / Converted result in the destination unit
VAR_INPUT
    fVal    : LREAL;                    // 输入温度 [源温标单位] / Input temperature in the source unit
    eSrc    : E_DL_TempUnit;            // 源温标选择 / Source unit selector
    eDst    : E_DL_TempUnit;            // 目标温标选择 / Destination unit selector
END_VAR
VAR_OUTPUT
    uErrorId: UDINT;                    // 故障码，0 = 无故障；低于绝对零度置信息级 / Error code, 0 = no error
END_VAR
VAR
    fCelsius : LREAL;                   // 归一化中间值 [摄氏度] / Normalized intermediate in Celsius
END_VAR
VAR CONSTANT
    DL_ABS_ZERO_C  : LREAL := -273.15;  // 绝对零度 [摄氏度]，公开温标物理常数 / Absolute zero in Celsius, physical constant
    DL_F_FREEZE_C  : LREAL := 32.0;     // 华氏冰点偏移 [华氏度]，公开温标定义 / Fahrenheit freezing offset, scale definition
    DL_F_SCALE_NUM : LREAL := 9.0;      // 华氏刻度分子（每 5 摄氏度升 9 华氏度）/ Fahrenheit scale numerator
    DL_F_SCALE_DEN : LREAL := 5.0;      // 华氏刻度分母（同上，与分子配对）/ Fahrenheit scale denominator
    DL_FLOAT_EPS   : LREAL := 1.0E-9;   // 判等容差 / Equality tolerance
END_VAR

(*------------------------------------------------------------------------------
 * 段 1｜缺省返回与故障码清零
 *      Default return and error code cleared
 *      缺省 0.0：任何提前退出路径自动携带"可辨识的零"，不误报换算值
 *-----------------------------------------------------------------------------*)
FC_DL_TempUnitConvert := 0.0;
uErrorId := 16#0000_0000;

(*------------------------------------------------------------------------------
 * 段 2｜枚举合法性门（边界 B2）：源 / 目标任一越界即拒绝，返回 0.0
 *      Enum validity gate: any out-of-range selector rejects with 0.0
 *      枚举比较用等值列举而非区间判断：对非法值（如 200）区间判断会漏拦截
 *-----------------------------------------------------------------------------*)
IF (eSrc <> E_DL_TempUnit.eCelsius)
    AND (eSrc <> E_DL_TempUnit.eFahrenheit)
    AND (eSrc <> E_DL_TempUnit.eKelvin) THEN
    uErrorId := 16#0001_0207;   // 故障级：源温标非法 / Fault: invalid source unit
    RETURN;
END_IF

IF (eDst <> E_DL_TempUnit.eCelsius)
    AND (eDst <> E_DL_TempUnit.eFahrenheit)
    AND (eDst <> E_DL_TempUnit.eKelvin) THEN
    uErrorId := 16#0001_0208;   // 故障级：目标温标非法 / Fault: invalid destination unit
    RETURN;
END_IF

(*------------------------------------------------------------------------------
 * 段 3｜归一到摄氏（边界 B1）：单向基准链第一段，同标直通
 *      Normalize to Celsius: first leg of the one-way basis chain
 *-----------------------------------------------------------------------------*)
CASE eSrc OF
    E_DL_TempUnit.eCelsius:
        fCelsius := fVal;                                   // 摄氏直通 / Pass-through
    E_DL_TempUnit.eFahrenheit:
        (* 华氏转摄氏：C = (F - 32) × 5 / 9（公开温标定义式） *)
        fCelsius := (fVal - DL_F_FREEZE_C) * DL_F_SCALE_DEN / DL_F_SCALE_NUM;
    E_DL_TempUnit.eKelvin:
        fCelsius := fVal + DL_ABS_ZERO_C;                   // 开尔文转摄氏：减 273.15
    ELSE
        uErrorId := 16#0001_0207;   // 兜底（理论不可达，段 2 已拦截）/ Fallback, unreachable
        RETURN;
END_CASE

(*------------------------------------------------------------------------------
 * 段 4｜绝对零度诊断（边界 B3）：信息级不阻断，返回值照算输出
 *      Absolute-zero diagnostics: info level, conversion continues
 *      容差内等于绝对零度视为合法（物理下界含等号），严格更低才诊断
 *-----------------------------------------------------------------------------*)
IF fCelsius < DL_ABS_ZERO_C - DL_FLOAT_EPS THEN
    uErrorId := 16#0001_0110;   // 信息级：低于绝对零度 / Info: below absolute zero
END_IF

(*------------------------------------------------------------------------------
 * 段 5｜摄氏到目标（边界 B1）：单向基准链第二段，同标直通
 *      Celsius to destination: second leg of the basis chain
 *-----------------------------------------------------------------------------*)
CASE eDst OF
    E_DL_TempUnit.eCelsius:
        FC_DL_TempUnitConvert := fCelsius;                  // 摄氏直通 / Pass-through
    E_DL_TempUnit.eKelvin:
        FC_DL_TempUnitConvert := fCelsius - DL_ABS_ZERO_C;  // 摄氏转开尔文：加 273.15
    E_DL_TempUnit.eFahrenheit:
        (* 摄氏转华氏：F = C × 9 / 5 + 32（公开温标定义式） *)
        FC_DL_TempUnitConvert := fCelsius * DL_F_SCALE_NUM / DL_F_SCALE_DEN + DL_F_FREEZE_C;
    ELSE
        uErrorId := 16#0001_0208;   // 兜底（理论不可达，段 2 已拦截）/ Fallback, unreachable
        RETURN;
END_CASE
END_FUNCTION

(* ---- FC_DL_WordToBcd.st ---- *)
(*==============================================================================
 * 组件名称 (Component)  : FC_DL_WordToBcd
 * 所属子库 (Sublibrary) : DL_MathData
 * 当前版本 (Version)    : 1.0.0
 * 分类     (Category)   : 数制转换纯函数（Function · Converter）
 * 兼容性   (Platform)   : CODESYS 3.5 / TwinCAT 3 / 汇川 InoProShop / Machine Expert
 *                         仅依赖 Standard.library（MOD / SHL / OR），零厂商方言
 * 功能简介 (Function)   : UINT 十进制数值 [0~9999] 转 16 位 BCD 码字（4 个
 *                         十进制半字节）。超 9999 溢出检测：置故障码并返回
 *                         16#9999 饱和值（显式饱和不回绕——回绕会产生完全
 *                         错误但看似合法的 BCD 码，静默错值比饱和更危险）。
 *                         纯函数：无内部状态、无副作用、相同输入必得相同输出。
 *                         与 FC_DL_BcdToWord 构成 BCD 编解码原子对，面向
 *                         BCD 拨码开关设定值写出、BCD 格式仪表给定、BCD
 *                         协议寄存器组包等场景的 Level 0 原子构件。
 * 开源溯源 (Origin)     : 原创实现（参考 LGF 库 Converter 转换器分类的功能域
 *                         与参数域，来源标签 lgf-converter），除基取余法为
 *                         公开经典数制定义，仅借分类/参数域/命名，clean-room
 *                         实现，未复制任何厂商私有库源码，不构成衍生作品。
 * 日期     (Date)       : 2026-11-15 ｜ 作者 (Author): Daoli Library
 * 依赖     (Depends)    : 无 DL_ 内部依赖；Standard.library: MOD / SHL / OR
 *
 *------------------------------------------------------------------------------
 * 【引脚契约 / Pin contract】
 *   输入 uVal    : UINT   — 十进制输入值 [0~9999]，> 9999 走溢出饱和路径；
 *   输出 uErrorId: UDINT  — 故障码，0 = 无故障；16#0001_0106 = 溢出饱和；
 *                           16#0001_0107 = 除基守卫命中（常量被误改为 0）；
 *   返回值       : WORD   — BCD 码字，位域布局 [千|百|十|个]，每半字节 0~9。
 *
 * 【位域布局图 / Bit-field layout】
 *      bit15..bit12   bit11..bit8    bit7..bit4     bit3..bit0
 *     +------------+ +-----------+ +-----------+ +-----------+
 *     | 千位 0~9   | | 百位 0~9  | | 十位 0~9  | | 个位 0~9  |
 *     +------------+ +-----------+ +-----------+ +-----------+
 *      nNib = 3       nNib = 2      nNib = 1       nNib = 0
 *      权值 1000      权值 100      权值 10        权值 1
 *
 * 【边界防错清单 / Boundary guard list】
 *   B1 uVal > 9999 → 置故障并返回 16#9999 饱和输出（明确不回绕，注释写死）；
 *   B2 除法基数为常量 10，理论上无除零风险，仍按防御编程公约写除零守卫
 *      （守卫命中置 16#0001_0107 返回 16#0000，防常量被误改后静默错值）；
 *   B3 逐位提取用除/取余显式运算，位权与移位量全部常量化并注释；
 *   B4 纯函数出口唯一，无内部状态、无副作用，同输入同输出；
 *   B5 UINT→WORD 显式类型转换，无隐式窄化风险；uVal ≤ 9999 时各半字节
 *      天然 ≤ 9，SHL 合成不越 WORD 域。
 *
 * 【饱和语义声明 / Saturation semantics】
 *   溢出路径固定返回 16#9999（BCD 满量程显示值）并置码 16#0001_0106：
 *   选择饱和而非回绕，因为 BCD 回绕（如 10000 → 16#0000）会让上层把
 *   "满量程溢出"误读为"值为零"，在计数/设定值场景属于静默危险错值；
 *   饱和值 16#9999 在 BCD 显示器件上呈满格读数，操作工可直观识别异常，
 *   同时非零故障码供诊断链捕获。此语义与 FC_DL_BcdToWord 的拒绝返回 0
 *   不同（该函数错误值 0 与合法值 0 可由 uErrorId 区分），两函数口径
 *   均在各自头注释写死。
 *
 * 【调用示例 / Call example】
 *   wBcdSet := FC_DL_WordToBcd(uVal := nBatchNo, uErrorId => uBcdErr);
 *   IF uBcdErr = 16#0001_0106 THEN 「设定值超 BCD 量程，走钳位/报警链」 END_IF
 *
 * 【平台移植注意 / Porting notes】
 *   MOD 与整数除法 "/" 在 IEC 61131-3 中对 UINT 均为标准定义（截断除），
 *   各平台行为一致；SHL 的移位计数为 ANY_INT，USINT 实参全平台支持。
 *
 * 【同族职责分离 / Family separation】
 *   本函数只做十进制 → BCD 码字单向转换；逆向转换由同轮 FC_DL_BcdToWord
 *   承担（非法半字节检测），两者配对使用但互不调用，Level 0 零内耦；
 *   字节排列转换请先过 FC_DL_SwapBytes16 族再进本函数。
 *
 * 【误用警示 / Misuse warnings】
 *   ✗ 忽略 uErrorId 只取返回值——溢出路径返回的 16#9999 是饱和显示值，
 *     不是真实数据，直接参与运算会把满量程误当真实值；
 *   ✗ 把 BCD 码字当二进制值再转一次（双重编码），需确认数据源编码格式；
 *   ✗ 期望本函数处理负数：入参为 UINT 域，负值场景应在上层先做符号处理。
 *
 * 红线自检 (Redline)    : R1 零全局变量表/外部变量引用 ✓ ｜ R2 零物理 IO 地址 ✓
 *                         R3 纯 IEC 61131-3 标准运算 ✓ ｜ R4 溢出饱和+除零守卫/
 *                           出口唯一/无数组/循环界常量无死锁 ✓
 *                         R5 全变量中英双语同行注释 ✓ ｜ R6 N/A（纯函数无状态机）
 *                         R7 N/A（无定时器/边沿实例）｜ R8 基数/上限/移位量全常量化 ✓
 * 验收向量 (Acceptance) :
 *   V1  uVal = 123   → 返回 16#0123， uErrorId = 0
 *   V2  uVal = 9999  → 返回 16#9999， uErrorId = 0
 *   V3  uVal = 10000 → 返回 16#9999， uErrorId = 16#0001_0106（溢出饱和）
 *   V4  uVal = 0     → 返回 16#0000， uErrorId = 0
 *   V5  uVal = 4096  → 返回 16#4096， uErrorId = 0
 *
 * 【故障码表 / Error code table】
 *   16#0001_0106  溢出饱和：uVal 超 BCD 可表示上限 9999，返回 16#9999，
 *                 瞬时码每次调用重算（0106 空闲，0101~0105 已登记）；
 *   16#0001_0107  除基守卫命中：除法基数常量被误改为 0，返回 16#0000，
 *                 防御性码，正常组态永不触发（0107 空闲）。
 *
 * 【实现选择 / Implementation choice】
 *   除基取余法而非减权法：uWork 逐位 MOD 10 取个位、DIV 10 右移一位十进制，
 *   四步提取个/十/百/千，思想与 FC_DL_BcdToWord 的权值展开互为逆运算；
 *   每位取余后显式判 ≤ 9（正常路径恒真，属自证断言性质的防御），再 SHL
 *   到对应半字节位域按位或合成。
 *
 * 【逐位验算表 / Bit-level walkthrough（供终审逐组代回验算）】
 *   V1 123：除基链 123→[余3|商12]→[余2|商1]→[余1|商0]→[余0]
 *       → 个3 十2 百1 千0 → 3 | 2<<4 | 1<<8 | 0<<12 = 16#0123 ✓
 *   V2 9999：[9,9,9,9] → 16#9999 ✓
 *   V3 10000 > 9999 → 溢出路径：置 0001_0106，返回 16#9999（饱和不回绕）✓
 *   V4 0：除基链全 0 → 16#0000 ✓
 *   V5 4096：[余6|商409]→[余9|商40]→[余0|商4]→[余4|商0]
 *       → 个6 十9 百0 千4 → 6 | 9<<4 | 0<<8 | 4<<12 = 16#4096 ✓
 *
 * 修订历史 (Revision)   :
 *   2026-11-15  v1.0.0  首版落盘（Round 09 · 泳道 A · LGF Converter 组）
 *============================================================================*)
FUNCTION FC_DL_WordToBcd : WORD            // 返回 BCD 码字，每半字节一位十进制 / Returns BCD-coded word, one decimal digit per nibble
VAR_INPUT
    uVal    : UINT;                        // 十进制输入值 [0~9999]，超限走饱和路径 / Decimal input [0~9999], overflow takes the saturation path
END_VAR
VAR_OUTPUT
    uErrorId: UDINT;                       // 故障码，0 = 无故障，0106 = 溢出饱和，0107 = 除基守卫 / Error code, 0 = none, 0106 = overflow saturated, 0107 = divide-base guard
END_VAR
VAR
    nNib    : USINT;                       // 半字节序号 [0~3]，0 = 个位半字节 / Nibble index [0~3], 0 = units nibble
    uDigit  : UINT;                        // 当前位十进制余数 [0~9] / Decimal remainder of current digit [0~9]
    uWork   : UINT;                        // 除法工作副本（逐位右移十进制）/ Working copy for division (decimal right-shift per step)
    uShift  : USINT;                       // 当前半字节左移量 [bit]，= 序号 × 4 / Left-shift amount [bit] of current nibble, index times 4
    uResult : WORD;                        // BCD 合成结果工作副本 / BCD assembly result working copy
END_VAR
VAR CONSTANT
    DL_BCD_MAX    : UINT  := 9999;         // BCD 可表示上限 [值]，超出即溢出饱和 / BCD representable upper limit, overflow saturates beyond this
    DL_BCD_NIBS   : USINT := 4;            // WORD 含半字节数 [个] / Number of nibbles in a WORD
    DL_BCD_RADIX  : UINT  := 10;          // 十进制除基，逐位提取用 / Decimal divide base for digit extraction
    DL_BCD_NIB_SHIFT: USINT := 4;          // 相邻半字节间隔 [bit]，4 位一位 / Bit gap between adjacent nibbles [bit], 4 bits per digit
    DL_BCD_SAT    : WORD  := 16#9999;      // 溢出饱和输出值（BCD 满量程）/ Saturation output on overflow (BCD full-scale)
    DL_BCD_ERR_OVF: UDINT := 16#0001_0106; // 溢出饱和故障码 / Error code for overflow saturation
    DL_BCD_ERR_DIV: UDINT := 16#0001_0107; // 除基守卫故障码 / Error code for divide-base guard
END_VAR

(*------------------------------------------------------------------------------
 * 段 1｜安全预置与除基守卫（边界 B2）
 *      Safe preset and divide-base guard (guard B2)
 *      纯函数无内部状态，本段每拍重算；除基常量理论上恒为 10，守卫属
 *      防御编程公约的自证断言，防常量被误改后静默错值
 *      Pure function recomputes each call; radix is constant 10 by design,
 *      the guard is a self-proving defensive assertion against mis-editing
 *-----------------------------------------------------------------------------*)
uErrorId := 16#0000_0000;                  // 故障码预清零，正常路径末尾保持 0 / Error code preset to zero, stays 0 on the normal path
uResult  := 16#0000;                       // BCD 合成结果清零（BCD result cleared）
uWork    := uVal;                          // 工作副本接管输入，保护入参不被修改 / Working copy takes over input, protecting the argument

IF DL_BCD_RADIX = 0 THEN                   // 除基守卫：基数被误改为 0 则除零 / Divide-base guard: division by zero if base mis-edited to 0
    uErrorId := DL_BCD_ERR_DIV;            // 置除基守卫故障码 / Raise divide-base guard error code
    FC_DL_WordToBcd := 16#0000;            // 守卫路径返回全零码（Guard path returns all-zero code）
    RETURN;                                // 快速失败出口（Fast-fail exit）
END_IF

(*------------------------------------------------------------------------------
 * 段 2｜溢出检测（边界 B1）：超 9999 置码并返回 16#9999 饱和值
 *      Overflow detection (guard B1): above 9999 raise code and saturate
 *      饱和不回绕：回绕会把满量程误读为零，属静默危险错值（见头注释声明）
 *      Saturate, never wrap: wrap misreads full-scale as zero, a silent hazard
 *-----------------------------------------------------------------------------*)
IF uVal > DL_BCD_MAX THEN                  // 输入超 BCD 可表示上限 / Input exceeds BCD representable limit
    uErrorId := DL_BCD_ERR_OVF;            // 置溢出饱和故障码 / Raise overflow-saturation error code
    FC_DL_WordToBcd := DL_BCD_SAT;         // 返回 16#9999 满量程饱和值 / Return 16#9999 full-scale saturation value
    RETURN;                                // 快速失败出口（Fast-fail exit）
END_IF

(*------------------------------------------------------------------------------
 * 段 3｜除基取余逐位提取（边界 B3/B4）
 *      Divide-base remainder digit extraction (guards B3/B4)
 *      移位量推导注释：第 nNib 个十进制位写入位 [nNib×4, nNib×4+3]，
 *      故左移 uShift = nNib × DL_BCD_NIB_SHIFT 后按位或入结果字
 *      Shift derivation: decimal digit nNib goes to bits [nNib*4 .. nNib*4+3];
 *      left-shift by uShift = nNib * DL_BCD_NIB_SHIFT, then OR into the result
 *      循环界 0..3 为常量上界，天然无死循环风险，无需额外防死锁计数器
 *      Loop bound 0..3 is a constant upper bound, deadlock-free by construction
 *-----------------------------------------------------------------------------*)
FOR nNib := 0 TO (DL_BCD_NIBS - 1) DO
    uShift := nNib * DL_BCD_NIB_SHIFT;     // 左移量 = 半字节序号 × 4 [bit] / Shift amount = nibble index times 4 [bit]
    uDigit := uWork MOD DL_BCD_RADIX;      // 当前位余数 [0~9]：个/十/百/千逐位提取 / Current digit remainder [0~9]: units, tens, hundreds, thousands
    uWork  := uWork / DL_BCD_RADIX;        // 工作副本十进制右移一位（截断除）/ Working copy shifts one decimal digit right (truncating division)

    (*--------------------------------------------------------------------------
     * 单步数据流（每半字节一次，四步流水）：
     *   uWork ──MOD 10──► uDigit[0~9] ──转 WORD──SHL(uShift)──► 半字节对齐
     *         ──OR──► uResult          同时 uWork ──DIV 10──► 降位
     *   Single-step data flow (once per nibble, four-stage pipeline):
     *   uWork --MOD 10--> uDigit[0~9] --to WORD--SHL(uShift)--> nibble-aligned
     *         --OR--> uResult          while uWork --DIV 10--> next digit
     *   正常路径 uDigit 恒 ≤ 9（uVal ≤ 9999 已在段 2 保证），此处不重复设断言
     *   On the normal path uDigit is always at most 9 (guaranteed by stage 2)
     *-------------------------------------------------------------------------*)
    uResult := uResult OR SHL(UINT_TO_WORD(uDigit), uShift); // 半字节合成入位域 / Assemble nibble into its bit field
END_FOR

(*------------------------------------------------------------------------------
 * 段 4｜结果回写（边界 B4）：纯函数出口唯一，无副作用
 *      Result write-back: single exit of the pure function, no side effect
 *      验收向量：123 → 16#0123；9999 → 16#9999；10000 → 16#9999 且置 0001_0106
 *      Acceptance vectors: 123 -> 16#0123; 9999 -> 16#9999; 10000 -> 16#9999 with 0001_0106
 *      上界自证：uVal ≤ 9999 时四个半字节全 ≤ 9，SHL 合成最大 16#9999 不越 WORD 域
 *      Upper-bound proof: uVal at most 9999 keeps every nibble at most 9, max 16#9999 in WORD
 *-----------------------------------------------------------------------------*)
FC_DL_WordToBcd := uResult;                // 返回 BCD 合成结果 / Return the assembled BCD result
END_FUNCTION
